TYPE "UDT_Service_Setup"
VERSION : 0.1
   STRUCT
      stepOrderOp : UInt;
      stepOrder { ExternalWritable := 'False'; S7_SetPoint := 'False'} : "UDT_Service_StepOrder";
      parameterIndexOp : UInt;
      parameterIndex { ExternalWritable := 'False'} : Byte;
   END_STRUCT;

END_TYPE

